(* IEC 61131-3 sources: llm-plc-st-eval/data/processed_definitivo/gpt-4o-2024-08-06/C4/few_shot, 3 files *)

(* ---- ejec_1.st ---- *)
FUNCTION_BLOCK FB_D
VAR_INPUT
    demanda : BOOL; (* Señal de demanda de operación *)
    falla1 : BOOL; (* Indica si la bomba 1 ha fallado *)
    falla2 : BOOL; (* Indica si la bomba 2 ha fallado *)
END_VAR
VAR_OUTPUT
    bomba1 : BOOL; (* Control de la bomba 1 *)
    bomba2 : BOOL; (* Control de la bomba 2 *)
    almFalla : BOOL; (* Alarma de falla de bomba *)
END_VAR
VAR
    turno : BOOL; (* Indica cuál bomba debe operar en el siguiente ciclo *)
    fDem : R_TRIG; (* Detector de flanco de subida para la señal de demanda *)
END_VAR

(* Detecta un flanco de subida en la señal de demanda *)
fDem(CLK := demanda);

(* Alterna el turno cada vez que hay un nuevo flanco de subida en la demanda *)
IF fDem.Q THEN
    turno := NOT turno;
END_IF

(* Lógica de control de bombas y manejo de fallas *)
IF demanda THEN
    IF turno THEN
        (* Si es el turno de la bomba 1 y no hay falla, activa bomba 1 *)
        bomba1 := NOT falla1;
        (* Si la bomba 1 falla, intenta activar la bomba 2 si no ha fallado *)
        bomba2 := falla1 AND NOT falla2;
        (* Activa la alarma si la bomba 1 falla *)
        almFalla := falla1;
    ELSE
        (* Si es el turno de la bomba 2 y no hay falla, activa bomba 2 *)
        bomba2 := NOT falla2;
        (* Si la bomba 2 falla, intenta activar la bomba 1 si no ha fallado *)
        bomba1 := falla2 AND NOT falla1;
        (* Activa la alarma si la bomba 2 falla *)
        almFalla := falla2;
    END_IF
ELSE
    (* Si no hay demanda, apaga ambas bombas y resetea la alarma *)
    bomba1 := FALSE;
    bomba2 := FALSE;
    almFalla := FALSE;
END_IF
END_FUNCTION_BLOCK

(* ---- ejec_2.st ---- *)
FUNCTION_BLOCK FB_D
VAR_INPUT
    demanda : BOOL; (* Señal de demanda para activar el sistema de bombeo *)
    falla1 : BOOL; (* Indica si hay una falla en la bomba 1 *)
    falla2 : BOOL; (* Indica si hay una falla en la bomba 2 *)
END_VAR
VAR_OUTPUT
    bomba1 : BOOL; (* Control de la bomba 1 *)
    bomba2 : BOOL; (* Control de la bomba 2 *)
    almFalla : BOOL; (* Alarma de falla si alguna bomba falla *)
END_VAR
VAR
    turno : BOOL; (* Variable para alternar entre las bombas *)
    fDem : R_TRIG; (* Detector de flanco de subida para la señal de demanda *)
END_VAR

(* Detecta un flanco de subida en la señal de demanda *)
fDem(CLK := demanda);

(* Si se detecta un nuevo flanco de subida en la demanda, alterna el turno *)
IF fDem.Q THEN
    turno := NOT turno;
END_IF

(* Lógica de control de bombas y alarma en función de la demanda y fallas *)
IF demanda THEN
    IF turno THEN
        (* Si es el turno de la bomba 1 y no hay falla, activa bomba 1 *)
        bomba1 := NOT falla1;
        (* Si hay falla en bomba 1, intenta activar bomba 2 si no está fallada *)
        bomba2 := falla1 AND NOT falla2;
        (* Activa la alarma si hay falla en bomba 1 *)
        almFalla := falla1;
    ELSE
        (* Si es el turno de la bomba 2 y no hay falla, activa bomba 2 *)
        bomba2 := NOT falla2;
        (* Si hay falla en bomba 2, intenta activar bomba 1 si no está fallada *)
        bomba1 := falla2 AND NOT falla1;
        (* Activa la alarma si hay falla en bomba 2 *)
        almFalla := falla2;
    END_IF
ELSE
    (* Si no hay demanda, apaga ambas bombas y resetea la alarma *)
    bomba1 := FALSE;
    bomba2 := FALSE;
    almFalla := FALSE;
END_IF
END_FUNCTION_BLOCK

(* ---- ejec_3.st ---- *)
FUNCTION_BLOCK FB_D
VAR_INPUT
    demanda : BOOL; (* Señal de demanda para activar las bombas *)
    falla1 : BOOL;  (* Indica si hay una falla en la bomba 1 *)
    falla2 : BOOL;  (* Indica si hay una falla en la bomba 2 *)
END_VAR
VAR_OUTPUT
    bomba1 : BOOL;  (* Estado de la bomba 1: activa o inactiva *)
    bomba2 : BOOL;  (* Estado de la bomba 2: activa o inactiva *)
    almFalla : BOOL; (* Alarma de falla en la bomba activa *)
END_VAR
VAR
    turno : BOOL;   (* Variable para alternar el uso de las bombas *)
    fDem : R_TRIG;  (* Detector de flanco ascendente para la demanda *)
END_VAR

(* Detecta el flanco ascendente de la señal de demanda *)
fDem(CLK := demanda);

(* Alterna el turno de las bombas en cada nueva demanda *)
IF fDem.Q THEN
    turno := NOT turno;
END_IF

(* Lógica de control de las bombas y alarmas *)
IF demanda THEN
    IF turno THEN
        (* Si es el turno de la bomba 1 *)
        bomba1 := NOT falla1; (* Activa bomba 1 si no hay falla *)
        bomba2 := falla1 AND NOT falla2; (* Activa bomba 2 si falla 1 y no falla 2 *)
        almFalla := falla1; (* Alarma si hay falla en bomba 1 *)
    ELSE
        (* Si es el turno de la bomba 2 *)
        bomba2 := NOT falla2; (* Activa bomba 2 si no hay falla *)
        bomba1 := falla2 AND NOT falla1; (* Activa bomba 1 si falla 2 y no falla 1 *)
        almFalla := falla2; (* Alarma si hay falla en bomba 2 *)
    END_IF
ELSE
    (* Si no hay demanda, ambas bombas y la alarma están inactivas *)
    bomba1 := FALSE;
    bomba2 := FALSE;
    almFalla := FALSE;
END_IF
END_FUNCTION_BLOCK
